(* Tests log record ownership and cloning. *)
FUNCTION_BLOCK FB_TestLogRecord EXTENDS FB_TestSuite
VAR_INPUT
END_VAR
VAR_OUTPUT
END_VAR
VAR
END_VAR

THIS^.testCloneToIsIndependent();

(* cloneTo deep copies a record, its resource, scope and every owned value, so a processor can keep the clone after the logger frees the source. Cloning into an assigned destination is refused so the existing record is not leaked. *)
METHOD testCloneToIsIndependent : REFERENCE TO FB_Test
VAR_INPUT
END_VAR
VAR
	resource: FB_Resource('resource.schema');
	provider: FB_LoggerProvider(resource);
	scope: FB_InstrumentationScope('scope.name', '1.0.0', 'scope.schema');
	logger: FB_Logger(scope, provider);
	timestamp: ULINT := 123456789;
	traceIdBytes: ARRAY [0..15] OF BYTE := [0, 1, 2, 3, 4, 5, 6, 7, 8, 9, 10, 11, 12, 13, 14, 15];
	spanIdBytes: ARRAY [0..7] OF BYTE := [16, 17, 18, 19, 20, 21, 22, 23];
	cloneSuccess: BOOL;
	cloneFailureResult: E_LogRecordCloneFailureReason;
	attributesSuccess: BOOL;
	attributesFailureReason: E_AttributesFailureReason;
	pClone: POINTER TO FB_LogRecord;
	pSourceResourceAttribute: POINTER TO FB_KeyValue;
	pClonedResourceAttribute: POINTER TO FB_KeyValue;
	pSourceScopeAttribute: POINTER TO FB_KeyValue;
	pClonedScopeAttribute: POINTER TO FB_KeyValue;
	pSourceRecordAttribute: POINTER TO FB_KeyValue;
	pClonedRecordAttribute: POINTER TO FB_KeyValue;
	pSourceString: POINTER TO FB_String;
	pClonedString: POINTER TO FB_String;
END_VAR
TcUnit.TEST('testCloneToIsIndependent');
	// Arrange: a source record with event name, body, IDs and one attribute at each level
	attributesSuccess := resource.attributes.setStringAttribute(
		key:='resource.key',
		value:='resource.value',
		failureReason=>attributesFailureReason
	);
	THIS^.AssertTrue(attributesSuccess, 'Expected resource attribute creation to succeed');
	attributesSuccess := scope.attributes.setStringAttribute(
		key:='scope.key',
		value:='scope.value',
		failureReason=>attributesFailureReason
	);
	THIS^.AssertTrue(attributesSuccess, 'Expected scope attribute creation to succeed');

	logger
		.startLogRecord(severityNumber:=E_SeverityNumber.INFO)
		.setTimestamp(timestamp)
		.setEventName('record.event')
		.setBody('record.body')
		._setTraceId(ADR(traceIdBytes), SIZEOF(traceIdBytes))
		._setSpanId(ADR(spanIdBytes), SIZEOF(spanIdBytes))
		._setFlags(16#01)  // sampled
		.setStringAttribute('record.key', 'record.value');
	THIS^.AssertTrue(logger.pLogRecord <> 0, 'Expected startLogRecord to build a source log record');

	// Clone: the first clone succeeds, a second into the same destination is refused
	IF logger.pLogRecord <> 0 THEN
		// no builder sets droppedAttributesCount; set by hand so the clone has a non-default value to copy
		logger.pLogRecord^.droppedAttributesCount := 4;
		cloneSuccess := logger.pLogRecord^.cloneTo(
			pDest:=pClone,
			failureReason=>cloneFailureResult
		);
		THIS^.AssertTrue(cloneSuccess, 'Expected log record clone to succeed');
		THIS^.AssertTrue(pClone <> 0, 'Expected a cloned log record');
		THIS^.AssertTrue(pClone <> logger.pLogRecord, 'Expected a distinct log record allocation');

		cloneSuccess := logger.pLogRecord^.cloneTo(
			pDest:=pClone,
			failureReason=>cloneFailureResult
		);
		THIS^.AssertFalse(cloneSuccess, 'Expected cloning into an assigned destination to fail');
		THIS^.AssertTrue(
			cloneFailureResult = E_LogRecordCloneFailureReason.DESTINATION_ALREADY_ASSIGNED,
			'Expected the DESTINATION_ALREADY_ASSIGNED reason when cloning into an assigned destination'
		);
	END_IF

	// Copied fields: equal values, distinct allocations for every owned value
	IF pClone <> 0 AND_THEN logger.pLogRecord <> 0 THEN
		THIS^.AssertTrue(pClone^.severityNumber = logger.pLogRecord^.severityNumber, 'Expected severity number to be cloned');
		THIS^.AssertTrue(pClone^.timestamp = logger.pLogRecord^.timestamp, 'Expected timestamp to be cloned');
		THIS^.AssertEquals_UDINT(logger.pLogRecord^.droppedAttributesCount, pClone^.droppedAttributesCount, 'Expected dropped record attribute count to be cloned');
		THIS^.AssertEquals_STRING(logger.pLogRecord^.resource.schemaUrl, pClone^.resource.schemaUrl, 'Expected resource schema URL to be cloned');
		THIS^.AssertEquals_UDINT(logger.pLogRecord^.resource.droppedAttributesCount, pClone^.resource.droppedAttributesCount, 'Expected dropped resource attribute count to be cloned');
		THIS^.AssertEquals_STRING(logger.pLogRecord^.scope.name, pClone^.scope.name, 'Expected scope name to be cloned');
		THIS^.AssertEquals_STRING(logger.pLogRecord^.scope.version, pClone^.scope.version, 'Expected scope version to be cloned');
		THIS^.AssertEquals_STRING(logger.pLogRecord^.scope.schemaUrl, pClone^.scope.schemaUrl, 'Expected scope schema URL to be cloned');
		THIS^.AssertEquals_UDINT(logger.pLogRecord^.scope.droppedAttributesCount, pClone^.scope.droppedAttributesCount, 'Expected dropped scope attribute count to be cloned');
		THIS^.AssertTrue(pClone^.eventName <> logger.pLogRecord^.eventName, 'Expected event name allocation to be cloned');
		THIS^.AssertTrue(pClone^.eventName^.pString <> logger.pLogRecord^.eventName^.pString, 'Expected event name string allocation to be cloned');
		THIS^.AssertEquals_STRING(logger.pLogRecord^.eventName^.pString^, pClone^.eventName^.pString^, 'Expected event name value to be cloned');
		THIS^.AssertTrue(pClone^.traceId <> logger.pLogRecord^.traceId, 'Expected trace ID allocation to be cloned');
		THIS^.AssertTrue(MEMCMP(ADR(pClone^.traceId^.bytes), ADR(logger.pLogRecord^.traceId^.bytes), SIZEOF(pClone^.traceId^.bytes)) = 0, 'Expected trace ID value to be cloned');
		THIS^.AssertEquals_UDINT(1, pClone^.flags, 'Expected the sampled trace flag to be cloned');
		THIS^.AssertTrue(pClone^.spanId <> logger.pLogRecord^.spanId, 'Expected span ID allocation to be cloned');
		THIS^.AssertTrue(MEMCMP(ADR(pClone^.spanId^.bytes), ADR(logger.pLogRecord^.spanId^.bytes), SIZEOF(pClone^.spanId^.bytes)) = 0, 'Expected span ID value to be cloned');
		THIS^.AssertTrue(pClone^.body <> logger.pLogRecord^.body, 'Expected body allocation to be cloned');
		pSourceString := logger.pLogRecord^.body;
		pClonedString := pClone^.body;
		THIS^.AssertTrue(pClonedString^.pString <> pSourceString^.pString, 'Expected body string allocation to be cloned');
		THIS^.AssertEquals_STRING(pSourceString^.pString^, pClonedString^.pString^, 'Expected body value to be cloned');

		// Attributes: each level's attribute, key and value are new allocations
		logger.pLogRecord^.resource.attributes.reset();
		pClone^.resource.attributes.reset();
		pSourceResourceAttribute := logger.pLogRecord^.resource.attributes.next();
		pClonedResourceAttribute := pClone^.resource.attributes.next();
		THIS^.AssertTrue(pSourceResourceAttribute <> 0, 'Expected the source record to have a resource attribute');
		THIS^.AssertTrue(pClonedResourceAttribute <> 0, 'Expected the cloned record to have a resource attribute');
		IF pSourceResourceAttribute <> 0 AND_THEN pClonedResourceAttribute <> 0 THEN
			THIS^.AssertTrue(pClonedResourceAttribute <> pSourceResourceAttribute, 'Expected resource attribute allocation to be cloned');
			THIS^.AssertTrue(pClonedResourceAttribute^.pKey <> pSourceResourceAttribute^.pKey, 'Expected resource attribute key allocation to be cloned');
			THIS^.AssertTrue(pClonedResourceAttribute^.pVal <> pSourceResourceAttribute^.pVal, 'Expected resource attribute value allocation to be cloned');
		END_IF

		logger.pLogRecord^.scope.attributes.reset();
		pClone^.scope.attributes.reset();
		pSourceScopeAttribute := logger.pLogRecord^.scope.attributes.next();
		pClonedScopeAttribute := pClone^.scope.attributes.next();
		THIS^.AssertTrue(pSourceScopeAttribute <> 0, 'Expected the source record to have a scope attribute');
		THIS^.AssertTrue(pClonedScopeAttribute <> 0, 'Expected the cloned record to have a scope attribute');
		IF pSourceScopeAttribute <> 0 AND_THEN pClonedScopeAttribute <> 0 THEN
			THIS^.AssertTrue(pClonedScopeAttribute <> pSourceScopeAttribute, 'Expected scope attribute allocation to be cloned');
			THIS^.AssertTrue(pClonedScopeAttribute^.pKey <> pSourceScopeAttribute^.pKey, 'Expected scope attribute key allocation to be cloned');
			THIS^.AssertTrue(pClonedScopeAttribute^.pVal <> pSourceScopeAttribute^.pVal, 'Expected scope attribute value allocation to be cloned');
		END_IF

		logger.pLogRecord^.attributes.reset();
		pClone^.attributes.reset();
		pSourceRecordAttribute := logger.pLogRecord^.attributes.next();
		pClonedRecordAttribute := pClone^.attributes.next();
		THIS^.AssertTrue(pSourceRecordAttribute <> 0, 'Expected the source record to have a record attribute');
		THIS^.AssertTrue(pClonedRecordAttribute <> 0, 'Expected the cloned record to have a record attribute');
		IF pSourceRecordAttribute <> 0 AND_THEN pClonedRecordAttribute <> 0 THEN
			THIS^.AssertTrue(pClonedRecordAttribute <> pSourceRecordAttribute, 'Expected record attribute allocation to be cloned');
			THIS^.AssertTrue(pClonedRecordAttribute^.pKey <> pSourceRecordAttribute^.pKey, 'Expected record attribute key allocation to be cloned');
			THIS^.AssertTrue(pClonedRecordAttribute^.pVal <> pSourceRecordAttribute^.pVal, 'Expected record attribute value allocation to be cloned');
		END_IF
	END_IF

	// Independence: the clone keeps its values after the logger frees the source
	logger.free();
	THIS^.AssertTrue(logger.pLogRecord = 0, 'Expected source log record to be deleted');

	IF pClone <> 0 THEN
		THIS^.AssertEquals_STRING('record.event', pClone^.eventName^.pString^, 'Expected cloned event name to survive source deletion');
		pClonedString := pClone^.body;
		THIS^.AssertEquals_STRING('record.body', pClonedString^.pString^, 'Expected cloned body to survive source deletion');
		THIS^.AssertEquals_UDINT(1, pClone^.resource.attributes.count, 'Expected cloned resource attributes to survive source deletion');
		THIS^.AssertEquals_UDINT(1, pClone^.scope.attributes.count, 'Expected cloned scope attributes to survive source deletion');
		THIS^.AssertEquals_UDINT(1, pClone^.attributes.count, 'Expected cloned record attributes to survive source deletion');
		pClone^.delete(pSelf:=pClone);
	END_IF
TcUnit.TEST_FINISHED();
END_METHOD

END_FUNCTION_BLOCK

(* stored: Version 1.1.0.1
   POU FB_TestLogRecord: Id {cf7b9e30-5700-468c-9441-fa4733ca3483}, SpecialFunc None
   Method testCloneToIsIndependent: Id {72ba3491-fa53-4815-8cd0-1a9a071d1081} *)
